(* IEC 61131-3 sources: SortJet_MasterSPS_Aufbau.fbsproj/09_Station/Stationen/Eckübergabe[204]/Aktionen, 3 files *)

(* ---- Eckuebergabe_Austransport_FB_V01_00_00.fb.st ---- *)
(* METADATA
{
	"v3Meta": {
		"objectGuid": "aec4a2b9-e42d-4dc6-88d8-ed1075e37aed"
	}
}
*)
FUNCTION_BLOCK Eckuebergabe_Austransport_FB_V01_00_00 EXTENDS Basic_Station_Austransport_FB_V01_00_00
VAR_IN_OUT

  // Anforderung an den Hubrahmen der Station
  blHubrahmenPositionieren : BOOL;
  elHubrahmenZielAchse     : Achsrichtung_EN;

END_VAR
VAR_INPUT

  // BOOL
  bpHubrahmenInPosition : BOOL; // Hubrahmen steht auf der angeforderten Achse

  // ENUM
  elAchseAustransport : Achsrichtung_EN; // Achse fuer den Austransport (Schnittstellendaten)

  // Bausteine
  Glastransport_X  : REFERENCE TO Eckuebergabe_Glastransport_FB_V01_00_00;
  Glastransport_Y  : REFERENCE TO Eckuebergabe_Glastransport_FB_V01_00_00;
  GlastransportAus : REFERENCE TO Eckuebergabe_Glastransport_FB_V01_00_00; // Austransport-Achse
  Hubrahmen        : REFERENCE TO ZylinderPneumatik_FB_V01_00_00;

END_VAR
//-------------------------------------------------------------------------------------------------
// AUSTRANSPORT
//-------------------------------------------------------------------------------------------------
IF ( BasisStationsParameter.bAustransport[wWand]
     AND bpAutomatikAktiv )
THEN

  // Ausnahmesituation
  IF ( Glastransport_X.bpFehler ) THEN
    Glastransport_X.bpAustransport             := FALSE;
    Glastransport_X.bpAustransportRueckwaertig := FALSE;
    BasisStationsParameter.wFehlerNummer := Glastransport_X.wpFehlerNr;
    steplAktion := STEP_900_E;
  END_IF

  IF ( Glastransport_Y.bpFehler ) THEN
    Glastransport_Y.bpAustransport             := FALSE;
    Glastransport_Y.bpAustransportRueckwaertig := FALSE;
    BasisStationsParameter.wFehlerNummer := Glastransport_Y.wpFehlerNr;
    steplAktion := STEP_900_E;
  END_IF

  IF ( Hubrahmen.bpFehler ) THEN
    blHubrahmenPositionieren := FALSE;
    BasisStationsParameter.awFehlerInformationen[1] := cZYLINDER_HUBRAHMEN;
    BasisStationsParameter.wFehlerNummer := Hubrahmen.wpFehlerNr;
    steplAktion := STEP_900_E;
  END_IF

  CASE steplAktion OF
    // AUSTRANSPORT =====================
    STEP_0_E:
      (* Hinweis:
         - Hubrahmen auf die Austransport-Achse stellen
      *)
      bpFehler := FALSE;

      elHubrahmenZielAchse     := elAchseAustransport;
      blHubrahmenPositionieren := TRUE;

      steplAktion := STEP_10_E;

    // AUSTRANSPORT =====================
    STEP_10_E:
      IF ( bpHubrahmenInPosition ) THEN
        blHubrahmenPositionieren := FALSE;

        steplAktion := STEP_100_E;
      END_IF

    // AUSTRANSPORT =====================
    STEP_100_E:
      (* Hinweis:
         - Austransport starten
      *)
      GlastransportAus.pAuftrag                   := BasisStationsParameter.pAuftrag[wWand];
      GlastransportAus.bpAustransport             := BasisStationsParameter.bAustransport[wWand] AND NOT BasisStationsParameter.bRueckwaertsTransportieren[wWand];
      GlastransportAus.bpAustransportRueckwaertig := BasisStationsParameter.bAustransport[wWand] AND     BasisStationsParameter.bRueckwaertsTransportieren[wWand];

      steplAktion := STEP_110_E;

    // AUSTRANSPORT =====================
    STEP_110_E:
      (* Hinweis:
         - Austransport abgeschlossen
      *)
      IF ( GlastransportAus.bpDone ) THEN
        GlastransportAus.bpAustransport             := FALSE;
        GlastransportAus.bpAustransportRueckwaertig := FALSE;

        steplAktion := STEP_1000_E;
      END_IF

    // AUSTRANSPORT =====================
    STEP_900_E:
      bpFehler := TRUE;
      BasisStationsParameter.bFehler := TRUE;

    // AUSTRANSPORT =====================
    STEP_1000_E:
      BasisStationsParameter.bAustransportAbgeschlossen[wWand] := TRUE;

  // AUSTRANSPORT =====================
  END_CASE
ELSE

  IF ( steplAktion > STEP_0_E ) THEN
    bpFehler := FALSE;
    BasisStationsParameter.bAustransportAbgeschlossen[wWand] := FALSE;

    Glastransport_X.bpAustransport             := FALSE;
    Glastransport_X.bpAustransportRueckwaertig := FALSE;
    Glastransport_Y.bpAustransport             := FALSE;
    Glastransport_Y.bpAustransportRueckwaertig := FALSE;
    blHubrahmenPositionieren                   := FALSE;

    steplAktion := STEP_0_E;
  END_IF

END_IF
END_FUNCTION_BLOCK

(* ---- Eckuebergabe_Eintransport_FB_V01_00_00.fb.st ---- *)
(* METADATA
{
	"v3Meta": {
		"objectGuid": "b3b83d22-15dc-44d1-82f1-6860a5f4b14c"
	}
}
*)
FUNCTION_BLOCK Eckuebergabe_Eintransport_FB_V01_00_00 EXTENDS Basic_Station_Eintransport_FB_V01_00_00
VAR_IN_OUT

  // Anforderung an den Hubrahmen der Station
  blHubrahmenPositionieren : BOOL;
  elHubrahmenZielAchse     : Achsrichtung_EN;

END_VAR
VAR_INPUT

  // BOOL
  bpHubrahmenInPosition : BOOL; // Hubrahmen steht auf der angeforderten Achse

  // ENUM
  elAchseEintransport : Achsrichtung_EN; // Achse des aktuellen Eintransports (Auftrag)
  elAchseAustransport : Achsrichtung_EN; // Achse fuer den Austransport (Schnittstellendaten)

  // Bausteine
  Glastransport_X  : REFERENCE TO Eckuebergabe_Glastransport_FB_V01_00_00;
  Glastransport_Y  : REFERENCE TO Eckuebergabe_Glastransport_FB_V01_00_00;
  GlastransportEin : REFERENCE TO Eckuebergabe_Glastransport_FB_V01_00_00; // Achse des aktuellen Eintransports
  GlastransportAus : REFERENCE TO Eckuebergabe_Glastransport_FB_V01_00_00; // Austransport-Achse
  Hubrahmen        : REFERENCE TO ZylinderPneumatik_FB_V01_00_00;

END_VAR
//-------------------------------------------------------------------------------------------------
// EINTRANSPORT
//-------------------------------------------------------------------------------------------------
IF ( BasisStationsParameter.bEintransport[wWand]
     AND bpAutomatikAktiv )
THEN

  // Ausnahmesituation
  IF ( Glastransport_X.bpFehler ) THEN
    Glastransport_X.bpEintransport             := FALSE;
    Glastransport_X.bpEintransportRueckwaertig := FALSE;
    Glastransport_X.bpVortransport             := FALSE;
    BasisStationsParameter.wFehlerNummer := Glastransport_X.wpFehlerNr;
    steplAktion := STEP_900_E;
  END_IF

  IF ( Glastransport_Y.bpFehler ) THEN
    Glastransport_Y.bpEintransport             := FALSE;
    Glastransport_Y.bpEintransportRueckwaertig := FALSE;
    Glastransport_Y.bpVortransport             := FALSE;
    BasisStationsParameter.wFehlerNummer := Glastransport_Y.wpFehlerNr;
    steplAktion := STEP_900_E;
  END_IF

  IF ( Hubrahmen.bpFehler ) THEN
    blHubrahmenPositionieren := FALSE;
    BasisStationsParameter.awFehlerInformationen[1] := cZYLINDER_HUBRAHMEN;
    BasisStationsParameter.wFehlerNummer := Hubrahmen.wpFehlerNr;
    steplAktion := STEP_900_E;
  END_IF

  CASE steplAktion OF
    // EINTRANSPORT =====================
    STEP_0_E:
      (* Hinweis:
         - Hubrahmen auf die Eintransport-Achse stellen
      *)
      bpFehler := FALSE;

      elHubrahmenZielAchse     := elAchseEintransport;
      blHubrahmenPositionieren := TRUE;

      steplAktion := STEP_10_E;

    // EINTRANSPORT =====================
    STEP_10_E:
      IF ( bpHubrahmenInPosition ) THEN
        blHubrahmenPositionieren := FALSE;

        steplAktion := STEP_100_E;
      END_IF

    // EINTRANSPORT =====================
    STEP_100_E:
      // ---------------------------------------------------------------------------------------
      //  STARTEN DES EINTRANSPORTS
      //
      //  Hinweis:
      //  - Eintransport ueber die Achse aus dem Auftrag
      // ---------------------------------------------------------------------------------------
      GlastransportEin.bpScheibentrennen          := BasisStationsParameter.bScheibentrennen[wWand];
      GlastransportEin.pAuftrag                   := BasisStationsParameter.pAuftrag[wWand];
      GlastransportEin.bpEintransport             := BasisStationsParameter.bEintransport[wWand] AND NOT BasisStationsParameter.bRueckwaertsTransportieren[wWand];
      GlastransportEin.bpEintransportRueckwaertig := BasisStationsParameter.bEintransport[wWand] AND     BasisStationsParameter.bRueckwaertsTransportieren[wWand];

      steplAktion := STEP_110_E;

    // EINTRANSPORT =====================
    STEP_110_E:
      IF ( GlastransportEin.bpDone ) THEN
        GlastransportEin.bpEintransport             := FALSE;
        GlastransportEin.bpEintransportRueckwaertig := FALSE;

        IF ( elAchseEintransport = elAchseAustransport ) THEN
          steplAktion := STEP_1000_E;
        ELSE
          steplAktion := STEP_200_E;
        END_IF
      END_IF

    // EINTRANSPORT =====================
    STEP_200_E:
      // ---------------------------------------------------------------------------------------
      //  UEBERGABE AN DIE AUSTRANSPORT-ACHSE
      //
      //  Hinweis:
      //  - Hubrahmen auf die Austransport-Achse stellen
      // ---------------------------------------------------------------------------------------
      elHubrahmenZielAchse     := elAchseAustransport;
      blHubrahmenPositionieren := TRUE;

      steplAktion := STEP_210_E;

    // EINTRANSPORT =====================
    STEP_210_E:
      IF ( bpHubrahmenInPosition ) THEN
        blHubrahmenPositionieren := FALSE;

        steplAktion := STEP_220_E;
      END_IF

    // EINTRANSPORT =====================
    STEP_220_E:
      (* Hinweis:
         - Austransport-Achse uebernimmt die Scheibe und faehrt sie auf den VorStop- Sensor
      *)
      GlastransportAus.pAuftrag       := BasisStationsParameter.pAuftrag[wWand];
      GlastransportAus.bpVortransport := TRUE;

      steplAktion := STEP_230_E;

    // EINTRANSPORT =====================
    STEP_230_E:
      IF ( GlastransportAus.bpDone ) THEN
        GlastransportAus.bpVortransport := FALSE;

        steplAktion := STEP_1000_E;
      END_IF

    // EINTRANSPORT =====================
    STEP_900_E:
      bpFehler := TRUE;
      BasisStationsParameter.bFehler := TRUE;

    // EINTRANSPORT =====================
    STEP_1000_E:
      BasisStationsParameter.bEintransportAbgeschlossen[wWand] := TRUE;

  // EINTRANSPORT =====================
  END_CASE
ELSE

  IF ( steplAktion > STEP_0_E ) THEN
    bpFehler := FALSE;
    BasisStationsParameter.bEintransportAbgeschlossen[wWand] := FALSE;

    Glastransport_X.bpEintransport             := FALSE;
    Glastransport_X.bpEintransportRueckwaertig := FALSE;
    Glastransport_X.bpVortransport             := FALSE;
    Glastransport_Y.bpEintransport             := FALSE;
    Glastransport_Y.bpEintransportRueckwaertig := FALSE;
    Glastransport_Y.bpVortransport             := FALSE;
    blHubrahmenPositionieren                   := FALSE;

    steplAktion := STEP_0_E;
  END_IF

END_IF
END_FUNCTION_BLOCK

(* ---- Eckuebergabe_Vortransport_FB_V01_00_00.fb.st ---- *)
(* METADATA
{
	"v3Meta": {
		"objectGuid": "516e6825-2e78-467d-914f-94fc332667ab"
	}
}
*)
FUNCTION_BLOCK Eckuebergabe_Vortransport_FB_V01_00_00 EXTENDS Basic_Station_Vortransport_FB_V01_00_00
VAR_IN_OUT

  // Anforderung an den Hubrahmen der Station
  blHubrahmenPositionieren : BOOL;
  elHubrahmenZielAchse     : Achsrichtung_EN;

END_VAR
VAR_INPUT

  // BOOL
  bpHubrahmenInPosition : BOOL; // Hubrahmen steht auf der angeforderten Achse

  // ENUM
  elAchseAustransport : Achsrichtung_EN; // Achse fuer den Austransport (Schnittstellendaten)

  // Bausteine
  Glastransport_X  : REFERENCE TO Eckuebergabe_Glastransport_FB_V01_00_00;
  Glastransport_Y  : REFERENCE TO Eckuebergabe_Glastransport_FB_V01_00_00;
  GlastransportAus : REFERENCE TO Eckuebergabe_Glastransport_FB_V01_00_00; // Austransport-Achse
  Hubrahmen        : REFERENCE TO ZylinderPneumatik_FB_V01_00_00;

END_VAR
//-------------------------------------------------------------------------------------------------
// VORTRANSPORT
//-------------------------------------------------------------------------------------------------
IF ( BasisStationsParameter.bVortransport[wWand]
     AND bpAutomatikAktiv )
THEN

  // Ausnahmesituation
  IF ( Glastransport_X.bpFehler ) THEN
    Glastransport_X.bpVortransport := FALSE;
    BasisStationsParameter.wFehlerNummer := Glastransport_X.wpFehlerNr;
    steplAktion := STEP_900_E;
  END_IF

  IF ( Glastransport_Y.bpFehler ) THEN
    Glastransport_Y.bpVortransport := FALSE;
    BasisStationsParameter.wFehlerNummer := Glastransport_Y.wpFehlerNr;
    steplAktion := STEP_900_E;
  END_IF

  IF ( Hubrahmen.bpFehler ) THEN
    blHubrahmenPositionieren := FALSE;
    BasisStationsParameter.awFehlerInformationen[1] := cZYLINDER_HUBRAHMEN;
    BasisStationsParameter.wFehlerNummer := Hubrahmen.wpFehlerNr;
    steplAktion := STEP_900_E;
  END_IF

  CASE steplAktion OF
    // VORTRANSPORT =====================
    STEP_0_E:
      (* Hinweis:
         - Hubrahmen auf die Austransport-Achse stellen
      *)
      bpFehler := FALSE;
      BasisStationsParameter.bVortransportAbgeschlossen[wWand] := FALSE;

      elHubrahmenZielAchse     := elAchseAustransport;
      blHubrahmenPositionieren := TRUE;

      steplAktion := STEP_10_E;

    // VORTRANSPORT =====================
    STEP_10_E:
      IF ( bpHubrahmenInPosition ) THEN
        blHubrahmenPositionieren := FALSE;

        steplAktion := STEP_100_E;
      END_IF

    // VORTRANSPORT =====================
    STEP_100_E:
      (* Hinweis:
         - Starten des Vortransports auf der Austransport-Achse
      *)
      GlastransportAus.bpVortransport := TRUE;

      steplAktion := STEP_110_E;

    // VORTRANSPORT =====================
    STEP_110_E:
      (* Hinweis:
         - Vortransport abgeschlossen
      *)
      IF ( GlastransportAus.bpDone ) THEN
        GlastransportAus.bpVortransport := FALSE;

        steplAktion := STEP_1000_E;
      END_IF

    // VORTRANSPORT =====================
    STEP_900_E:
      bpFehler := TRUE;
      BasisStationsParameter.bFehler := TRUE;

    // VORTRANSPORT =====================
    STEP_1000_E:
      BasisStationsParameter.bVortransportAbgeschlossen[wWand] := TRUE;

  // VORTRANSPORT =====================
  END_CASE
ELSE

  IF ( steplAktion > STEP_0_E ) THEN
    bpFehler := FALSE;
    BasisStationsParameter.bVortransportAbgeschlossen[wWand] := FALSE;

    Glastransport_X.bpVortransport := FALSE;
    Glastransport_Y.bpVortransport := FALSE;
    blHubrahmenPositionieren       := FALSE;

    steplAktion := STEP_0_E;
  END_IF

END_IF
END_FUNCTION_BLOCK
